Fanuc KAREL source: kt00552.KL

-- PROVISIONAL review KL for V770-1; original PC SHA256 c67c3f93274a2d54c4b7980c0110291d9e4431f52ea25a6fdfb3f2600388215f
-- Incomplete behavior may be omitted. Consult companion uncertainty JSON. Do not deploy.
PROGRAM KT00552
%NOLOCKGROUP
-- UNRESOLVED_DECL P1 type=000199
-- UNRESOLVED_DECL P2 type=000199
-- UNRESOLVED_DECL OUT type=000199
BEGIN
  -- UNRESOLVED_PC offsets 5-44; opcodes 49,7E,49,7E,60,7E,4A
  -- UNRESOLVED_PC offsets 49-53; opcodes 7F
END KT00552
